PROGRAM main
  VAR
    MARCHA AT %IX0.0  : BOOL; (* S1, pulsador NA *)
    PARADA AT %IX0.1  : BOOL; (* S2, pulsador NC: activa en reposo *)
    TERMICO AT %IX0.2 : BOOL; (* F1, contacto 95-96 NC: activo si no hay falla *)
    KM1 AT %QX0.0     : BOOL; (* contactor del motor *)
    H1 AT %QX0.1      : BOOL; (* piloto de falla *)
    H2 AT %QX0.2      : BOOL; (* piloto de marcha *)
  END_VAR
  VAR  (* added by the conversion: wires and edge detectors of the diagram *)
    _OR2_OUT : BOOL;
    _AND1_OUT : BOOL;
    _NOT10_OUT : BOOL;
  END_VAR

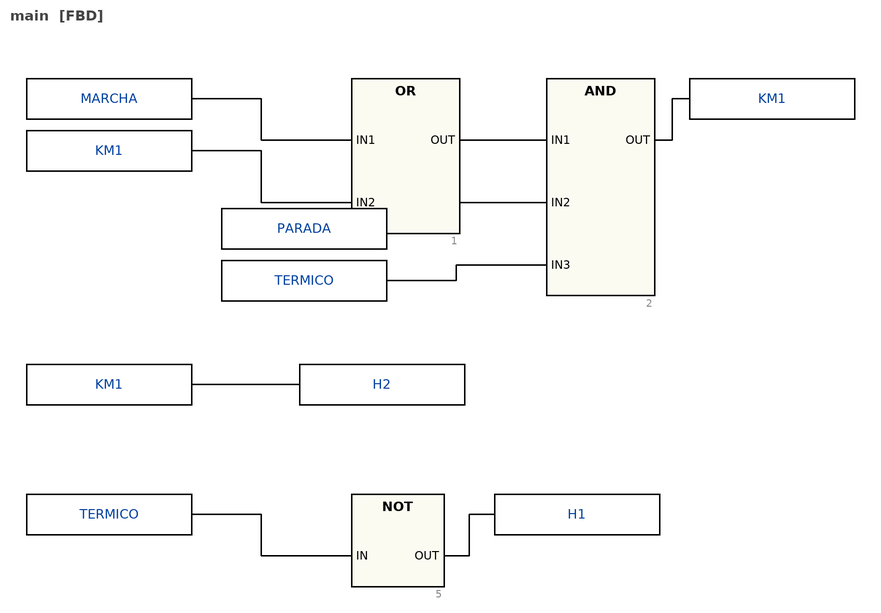
(* FBD diagram, written out as Structured Text *)
_OR2_OUT := MARCHA OR KM1;
_AND1_OUT := _OR2_OUT AND PARADA AND TERMICO;
KM1 := _AND1_OUT;
H2 := KM1;
_NOT10_OUT := NOT TERMICO;
H1 := _NOT10_OUT;
END_PROGRAM
